// TIA Portal V20 export
Screen "Pop-up_StyleConfigMESDownload"  654x462
